SUBAPPLICATION mapping_Softkeys (* Subapplication Type *)
  (* Standard: 61499-2 *)
  (* Version 1.0, 2023-01-29, Franz *)
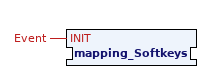
  EVENT_INPUT
    INIT;
  END_EVENT
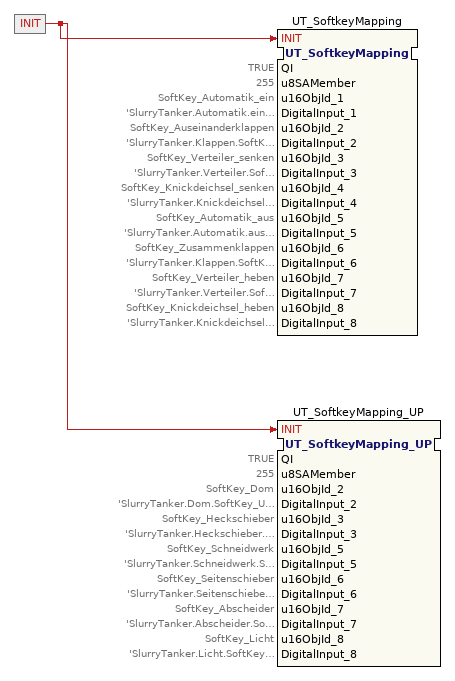
  FBS
    UT_SoftkeyMapping : UT_SoftkeyMapping(QI := TRUE, u8SAMember := 255, u16ObjId_1 := SoftKey_Automatik_ein, DigitalInput_1 := 'SlurryTanker.Automatik.ein.SoftKey', u16ObjId_2 := SoftKey_Auseinanderklappen, DigitalInput_2 := 'SlurryTanker.Klappen.SoftKey_heben.SoftKey', u16ObjId_3 := SoftKey_Verteiler_senken, DigitalInput_3 := 'SlurryTanker.Verteiler.SoftKey_senken.SoftKey', u16ObjId_4 := SoftKey_Knickdeichsel_senken, DigitalInput_4 := 'SlurryTanker.Knickdeichsel.SoftKey_senken.SoftKey', u16ObjId_5 := SoftKey_Automatik_aus, DigitalInput_5 := 'SlurryTanker.Automatik.aus.SoftKey', u16ObjId_6 := SoftKey_Zusammenklappen, DigitalInput_6 := 'SlurryTanker.Klappen.SoftKey_senken.SoftKey', u16ObjId_7 := SoftKey_Verteiler_heben, DigitalInput_7 := 'SlurryTanker.Verteiler.SoftKey_heben.SoftKey', u16ObjId_8 := SoftKey_Knickdeichsel_heben, DigitalInput_8 := 'SlurryTanker.Knickdeichsel.SoftKey_heben.SoftKey');
    UT_SoftkeyMapping_UP : UT_SoftkeyMapping_UP(QI := TRUE, u8SAMember := 255, u16ObjId_2 := SoftKey_Dom, DigitalInput_2 := 'SlurryTanker.Dom.SoftKey_UP.SoftKey', u16ObjId_3 := SoftKey_Heckschieber, DigitalInput_3 := 'SlurryTanker.Heckschieber.SoftKey_UP.SoftKey', u16ObjId_5 := SoftKey_Schneidwerk, DigitalInput_5 := 'SlurryTanker.Schneidwerk.SoftKey_UP.SoftKey', u16ObjId_6 := SoftKey_Seitenschieber, DigitalInput_6 := 'SlurryTanker.Seitenschieber.SoftKey_UP.SoftKey', u16ObjId_7 := SoftKey_Abscheider, DigitalInput_7 := 'SlurryTanker.Abscheider.SoftKey_UP.SoftKey', u16ObjId_8 := SoftKey_Licht, DigitalInput_8 := 'SlurryTanker.Licht.SoftKey_UP.SoftKey');
  END_FBS
  EVENT_CONNECTIONS
    INIT TO UT_SoftkeyMapping.INIT;
    INIT TO UT_SoftkeyMapping_UP.INIT;
  END_CONNECTIONS
END_SUBAPPLICATION
